Staubli VAL3: main.pgx

program main()
begin
  close(tCurrentTool)
  pPointRs.config.shoulder = lefty
  pPointRs2.config.shoulder = lefty
  mCurrentSpeed.tvel = 100.00
  mCurrentSpeed.blend = joint
  mCurrentSpeed.reach = 0.010
  mCurrentSpeed.leave = 0.010
  // Program PrecProg start
  // Program generated by RoboDK v6.0.7 for Staubli TS20 FL 100 TC on XX/XX/XXXX 18:00:00
  // Using nominal kinematics.
  call MoveJoint(12.34560,-45.67890,78.90130,-0.50000)
  call MoveLine(-640.585,506.981,371.534,136.641,31.137,-130.569)
  call MoveLine(0.500,-0.500,0.250,-180.000,0.005,-0.005)
  call MoveJoint(-12.34540,45.67850,-78.90000,0.50000)
  call MoveJoint(-12.34540,45.67850,-78.90000,0.50000)
  mCurrentSpeed.tvel = 66.667
  delay(0.002)
  delay(1.000)
  call MoveLine(-353.026,-90.135,331.702,164.619,39.324,-168.579)

  waitEndMove()
  // Program PrecProg end

end
